FUNCTION F_AnalogToEngUnit : LREAL
VAR_INPUT
	inpRawSignal	:	LREAL;
	IO_min			:	LREAL;
	IO_max			: 	LREAL;
	engMin			:   LREAL;
	engMax			:	LREAL;
END_VAR

F_AnalogToEngUnit	:= engMin + (inpRawSignal - IO_min) * ((engmax - engmin) / (IO_max - IO_min));

END_FUNCTION

(* stored: Version 1.1.0.1
   POU F_AnalogToEngUnit: Id {754c32c2-8cb1-4acd-8139-f0ef6fb6f60e}, SpecialFunc None *)
